FUNCTION_BLOCK FB_STOEBERSDS_MC_Power
(*

The function block used to activates software enable for an axis

Constructor: 		Patryk Panylo
Company:		E. Riexinger GmbH
Date:			22.09.2015
Version:			1.00

Date:			Revision:		Who:				Comment

*)
VAR_INPUT
	(* Input variables / Eingang Variablen *)
	bEnable						:BOOL;			(* Signal FB enable *)
	bRegulatorOn				:BOOL;			(* Enable the power stage *)
	bEnablePositive				:BOOL;			(* Advance movement enable in positive direction. *)
	bEnableNegative				:BOOL;			(* Advance movement enable in negative direction. *)
	lrOverride					:LREAL;			(* Velocity override in % for all motion commands. (0 <= Override <= 100.0) *)
END_VAR
VAR_OUTPUT
	(* Output variables / Ausgang Variablen *)
	bStatus						:BOOL;			(* Status = TRUE indicates that the axis is ready for operation. *)
	bError						:BOOL;			(* Error *)
	udnErrorNo					:UDINT;			(* Error number *)
	sErrorMsg					:STRING; 		(* Error message *)
END_VAR
VAR_IN_OUT
	(* Input Output variables / Ausgang Variablen *)
	Axis							:ST_AXIS_REF;
END_VAR
VAR
	(* Enummerations *)

	(* Variables *)
	tStatusDelay 					:TIME := t#300ms;

	(* References *)

	(* Interfaces *)

	(* Instances *)
	tonStatusDelay				:TON;
END_VAR


IF NOT bEnable
THEN
	Axis.stPlcToNc.stBaseDevice.bEnable := FALSE;                   		 (* Switch off *)
	tonStatusDelay(IN := FALSE,
				    PT := tStatusDelay);
ELSE

	IF NOT bRegulatorOn
	     OR Axis.stNcToPlc.stBaseDevice.bError
	THEN
		Axis.stPlcToNc.stBaseDevice.bEnable := FALSE;			(* Switch off *)
	ELSE
		Axis.stPlcToNc.stBaseDevice.bEnable := TRUE;                     	(* Switch on *)
	END_IF;

END_IF;

Axis.stPlcToNc.stBaseDevice.bFeedEnablePlus := bEnablePositive;
Axis.stPlcToNc.stBaseDevice.bFeedEnableMinus := bEnableNegative;

Axis.stPlcToNc.stBaseDevice.stCommandPositioning.nOverride := LREAL_TO_INT(lrOverride * 32767 / 200);

tonStatusDelay(IN := Axis.stNcToPlc.stBaseDevice.bEnabled,		(* Control enabled *)
			   PT := tStatusDelay);
bStatus := tonStatusDelay.Q;

bError := Axis.stNcToPlc.stBaseDevice.bError;                     (* Error *)

END_FUNCTION_BLOCK

(* stored: Version 1.1.0.1, ProductVersion 3.1.4024.15
   POU FB_STOEBERSDS_MC_Power: Id {626bb414-59c2-4a09-91a1-4c296bcb374a}, SpecialFunc None *)
